(* IEC 61131-3 sources: RootPLC/conformance/cases/codegen, 2 files *)

(* ---- ok_build_c_subset.st ---- *)
(* spec: [build.c.command] [build.c.file] [build.c.semantics] [build.c.faults] [build.c.subset] [build.c.oop]
   expect: ok
   run: PRG_Main cycles=5
   assert: n = 5
   assert: wrapped = -32768
   assert: rounded = 3
   assert: total = 15
   assert: avg > 2.99 AND avg < 3.01 *)
(* The v0 subset of the C back end in one program; the driver test
   tests/codegen_c.rs translates it to C, compiles it and compares every
   variable with the VM (with the clock advancing 10 ms per cycle, so the
   timer and counter also run there; the conformance runner does not
   advance the clock). *)
TYPE E_Mode : (IDLE, RUN, DONE); END_TYPE
TYPE ST_Stat : STRUCT
    count : INT;
    sum : DINT;
END_STRUCT; END_TYPE
TYPE T_Pct : INT (0..100); END_TYPE

FUNCTION Average : REAL
VAR_INPUT
    sum : DINT;
    count : INT := 1;
END_VAR
IF count = 0 THEN
    Average := 0.0;
ELSE
    Average := DINT_TO_REAL(sum) / INT_TO_REAL(count);
END_IF;
END_FUNCTION

FUNCTION_BLOCK FB_Acc
VAR_INPUT x : INT; END_VAR
VAR_OUTPUT stat : ST_Stat; END_VAR
stat.count := stat.count + 1;
stat.sum := stat.sum + x;
END_FUNCTION_BLOCK

PROGRAM PRG_Main
VAR
    n : INT;
    mode : E_Mode := E_Mode#IDLE;
    acc : FB_Acc;
    hist : ARRAY[1..5] OF INT;
    total : DINT;
    avg : REAL;
    wrapped : INT := 32767;
    rounded : DINT;
    pct : T_Pct := 50;
    pulses : CTU;
    blink : TON;
    k : INT;
END_VAR
n := n + 1;
hist[n] := n;
acc(x := n);
total := 0;
FOR k := 1 TO 5 DO
    IF hist[k] = 0 THEN
        CONTINUE;
    END_IF;
    total := total + hist[k];
END_FOR;
avg := Average(sum := acc.stat.sum, count := acc.stat.count);
CASE n OF
    1: mode := E_Mode#RUN;
    2..4: pct := pct + 10;
ELSE
    mode := E_Mode#DONE;
END_CASE;
IF n = 5 THEN
    wrapped := wrapped + 1;
    rounded := REAL_TO_DINT(2.5);
END_IF;
blink(IN := NOT blink.Q, PT := T#20ms);
pulses(CU := blink.Q, PV := 10);
END_PROGRAM

(* ---- ok_build_c_strings.st ---- *)
(* spec: [build.c.semantics] [build.c.strings] [build.c.subset]
   expect: ok
   run: PRG_Main cycles=2
   assert: short = 'abcde'
   assert: joined = 'ab-cd-ef'
   assert: n = 8
   assert: pos = 3
   assert: none = 0
   assert: empty_at = 1
   assert: l = 'ab'
   assert: r = 'ef'
   assert: m = 'cd'
   assert: m0 = 'ab'
   assert: ins = 'XYab-cd-ef'
   assert: ins_end = 'ab-cd-efXY'
   assert: del = 'ab-ef'
   assert: rep = 'ab-ZZZ-ef'
   assert: num = -42
   assert: bad = 0
   assert: neg = '-17'
   assert: dur = 'T#1m30s250ms'
   assert: zero = 'T#0ms'
   assert: yes = 'TRUE'
   assert: less
   assert: count = 2
   assert: r1 = '0.1'
   assert: r2 = '1E-5'
   assert: r3 = '1.5E16'
   assert: r4 = '100.0'
   assert: r5 = '-0.00025'
   assert: r6 = '0.0001'
   assert: d1 = 'D#2026-11-07'
   assert: t1 = 'TOD#12:30:15.25'
   assert: dt1 = 'DT#2026-11-07-08:09:10' *)
(* String functions at their edges, for the C back end; the driver test
   compares every variable with the VM. *)
PROGRAM PRG_Main
VAR
    short : STRING[5];
    joined : STRING;
    n : INT;
    pos : INT;
    none : INT;
    empty_at : INT;
    l, r, m, m0 : STRING;
    ins, ins_end, del, rep : STRING;
    num : INT;
    bad : INT;
    neg : STRING;
    dur : STRING;
    zero : STRING;
    yes : STRING;
    less : BOOL;
    count : INT;
    r1, r2, r3, r4, r5, r6 : STRING;
    d1, t1, dt1 : STRING;
END_VAR
count := count + 1;
short := CONCAT('abcd', 'efgh');
joined := CONCAT('ab', '-cd', '-ef');
n := LEN(joined);
pos := FIND(joined, '-');
none := FIND(joined, 'zz');
empty_at := FIND(joined, '');
l := LEFT(joined, 2);
r := RIGHT(joined, 2);
m := MID(joined, 2, 4);
m0 := MID(joined, 2, 0);
ins := INSERT(joined, 'XY', 0);
ins_end := INSERT(joined, 'XY', 99);
del := DELETE(joined, 3, 3);
rep := REPLACE(joined, 'ZZZ', 2, 4);
num := STRING_TO_INT('  -42 ');
bad := STRING_TO_INT('4x2');
neg := INT_TO_STRING(-17);
dur := TIME_TO_STRING(T#90s250ms);
zero := TIME_TO_STRING(T#0s);
yes := BOOL_TO_STRING(TRUE);
less := 'abc' < 'abd' AND 'ab' < 'abc' AND NOT ('b' < 'abc');
r1 := REAL_TO_STRING(0.1);
r2 := REAL_TO_STRING(1.0E-5);
r3 := REAL_TO_STRING(1.5E16);
r4 := REAL_TO_STRING(100.0);
r5 := LREAL_TO_STRING(-2.5E-4);
r6 := LREAL_TO_STRING(1.0E-4);
d1 := DATE_TO_STRING(D#2026-11-07);
t1 := TOD_TO_STRING(TOD#12:30:15.25);
dt1 := DT_TO_STRING(DT#2026-11-07-08:09:10);
END_PROGRAM
